(* CODESYS project SysParFeedRobot.xml

Project tree, tasks and I/O mapping:
  visualisation SysParFeedRobot
*)

// /SysParFeedRobot
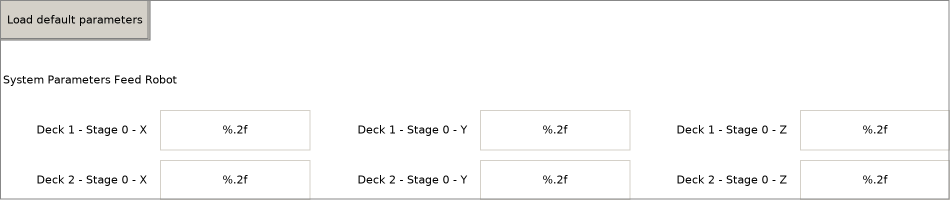
VISUALIZATION SysParFeedRobot  // 950x200
    Button (0,0 150x40), "Load default parameters"
        tap PRG_VisuTask_10ms._fbParametersCtrl._btnLoadDefaultParameters.xbtn
    Label (0,60 300x40), "System Parameters Feed Robot"
    Label (0,110 150x40), "Deck 1 - Stage 0 - X"
    Textfield (160,110 150x40), "%.2f", text variable: PersistentVars.scFeedrobot.RobotArm.DeckPositions[1].posX
        OnMouseUp: write the text variable via Default, min -25, max 25
    Label (320,110 150x40), "Deck 1 - Stage 0 - Y"
    Textfield (480,110 150x40), "%.2f", text variable: PersistentVars.scFeedrobot.RobotArm.DeckPositions[1].posY
        OnMouseUp: write the text variable via Default, min -25, max 25
    Label (640,110 150x40), "Deck 1 - Stage 0 - Z"
    Textfield (800,110 150x40), "%.2f", text variable: PersistentVars.scFeedrobot.RobotArm.DeckPositions[1].posZ
        OnMouseUp: write the text variable via Default, min 0, max 50
    Label (0,160 150x40), "Deck 2 - Stage 0 - X"
    Textfield (160,160 150x40), "%.2f", text variable: PersistentVars.scFeedrobot.RobotArm.DeckPositions[2].posX
        OnMouseUp: write the text variable via Default, min -25, max 25
    Label (320,160 150x40), "Deck 2 - Stage 0 - Y"
    Textfield (480,160 150x40), "%.2f", text variable: PersistentVars.scFeedrobot.RobotArm.DeckPositions[2].posY
        OnMouseUp: write the text variable via Default, min -25, max 25
    Label (640,160 150x40), "Deck 2 - Stage 0 - Z"
    Textfield (800,160 150x40), "%.2f", text variable: PersistentVars.scFeedrobot.RobotArm.DeckPositions[2].posZ
        OnMouseUp: write the text variable via Default, min 0, max 50
END_VISUALIZATION
